(* IEC 61131-3 sources: volt/packages/volt-lsp-iec/test-corpus/lenze-mid/Device/Plc Logic/Application/Library Manager/L_OEEA_BaseDependency, 3.26.4.8 (Lenze), 88 files *)

(* ---- ENUMOEECALCULATIONMODE.dut ---- *)
TYPE ENUMOEECALCULATIONMODE :
(
	STANDARD := 0,
	PART_SUMMERY := 1
);
END_TYPE

(* ---- ENUMOEEPARTTARGETMODE.dut ---- *)
TYPE ENUMOEEPARTTARGETMODE :
(
	SHIFTPARTTARGET := 0,
	PRODUCTPARTTARGET := 1
);
END_TYPE

(* ---- ENUMRUNRATEFREQUENCE.dut ---- *)
TYPE ENUMRUNRATEFREQUENCE :
(
	HOUR_1X := 1,
	HOUR_2X := 2,
	HOUR_4X := 4
);
END_TYPE

(* ---- ENUMSHIFTMODE.dut ---- *)
TYPE ENUMSHIFTMODE :
(
	SHIFT := 0,
	HOURS24 := 1,
	NOSCHEDULE := 2,
	SHIFT7DAYS := 3,
	HOURS24_7DAYS := 4
);
END_TYPE

(* ---- RT_DOWNTIME.dut ---- *)
TYPE RT_DOWNTIME :
STRUCT
	PARA : ARRAY [0..19] OF sc_RT_Downtime;
END_STRUCT
END_TYPE

(* ---- RT_STATUS_STRUCT.dut ---- *)
TYPE RT_STATUS_STRUCT :
STRUCT
	STATIONID : DINT;
	PARTID : DINT;
	TOTALPARTSOK : DINT;
	TOTALPARTSNOK : DINT;
	TOTALPARTSOK_2 : DINT;
	TOTALPARTSNOK_2 : DINT;
	PARTTYPEID : DINT;
	PARTTYPESTR : STRING(100);
	PRODMODE : INT;
	PRODMODESTR : STRING;
	PARTCYCLETIME : REAL;
	OPCYCLETIME : REAL;
	ALIVECOUNTER : DINT;
	ERROR : BOOL;
	WARNING : BOOL;
	DOWNTIMECODE : INT;
	SDOWNTIMESTR : STRING;
	REASONCODE : DINT;
	REASONCODESTR : STRING;
	DOWNTIMEACTIVE : BOOL;
END_STRUCT
END_TYPE

(* ---- RT_TIMER.dut ---- *)
TYPE RT_TIMER :
STRUCT
	TOK_PART : TIME;
	TNOK_PART : TIME;
	TOK_PART2 : TIME;
	TNOK_PART2 : TIME;
	TALIVECOUNTER : TIME;
	TERROR : ARRAY [0..19] OF TIME;
	TERRORDURATION : ARRAY [0..19] OF TIME;
	TWARNING : TIME;
	TWARNINGDURATION : TIME;
	TPARTTYPECHANGE : TIME;
	TPARTCYCLETIME : TIME;
	TOPCYCLETIME : TIME;
END_STRUCT
END_TYPE

(* ---- SC_RT_DOWNTIME.dut ---- *)
TYPE SC_RT_DOWNTIME :
STRUCT
	PRODUCTIONMODE : INT;
	DOWNTIMECODE : INT;
	REASONCODE : DINT;
	SREASONCODESTR : STRING;
END_STRUCT
END_TYPE

(* ---- SCACCESSPOINTS.dut ---- *)
TYPE SCACCESSPOINTS :
STRUCT
	TACTUALPLANNEDPRODUCTION : TIME;
	TSHIFTPLANNEDPRODUCTION : TIME;
	TACTUALALLTIME : TIME;
	TACTUALRUNTIME : TIME;
	TDOWNTIME : TIME;
	TORGDOWNTIME : TIME;
	TNONPRODUCTIVETIME : TIME;
	DIACTUALALLTIME : DINT;
	DIACTUALPLANNEDPRODUCTION : DINT;
	DISHIFTPLANNEDPRODUCTION : DINT;
	DIACTUALRUNTIME : DINT;
	DIDOWNTIME : DINT;
	DIORGDOWNTIME : DINT;
	DINONPRODUCTIVETIME : DINT;
	LRPARTSUMMERY : LREAL;
	LRACTUALPARTCOUNT : LREAL;
	RINCONSISTENTPARTCOUNTDEVIATION : REAL;
	XPRODUCTIONTARGETREACHED : BOOL;
	XCHANGEOVERTIMEACTIVE : BOOL;
	XCHANGEOVERTIMEEXCEEDED : BOOL;
END_STRUCT
END_TYPE

(* ---- SCACTUALPRODUCTION.dut ---- *)
TYPE SCACTUALPRODUCTION :
STRUCT
	XPRODUCTIONACTIVE : BOOL;
	XPRODUCTIONHOLD : BOOL;
	EOEECALCMODE : enumOEECalculationMode;
	EOEEPARTTARGETMODE : enumOEEPartTargetMode;
	IOEEKPIDECIMALS : INT := 1;
	RSETSPEEDVALUE : REAL;
	RSETSPEEDPERCENT : REAL;
	ITRIGGER : INT;
END_STRUCT
END_TYPE

(* ---- SCBATCH.dut ---- *)
TYPE SCBATCH :
STRUCT
	DIID : DINT;
	DIJOBID : DINT;
	SJOBNO : STRING;
	DIJOBTARGET : DINT;
END_STRUCT
END_TYPE

(* ---- SCBATCHPRODUCTEND.dut ---- *)
TYPE SCBATCHPRODUCTEND :
STRUCT
	XONBATCHIDCHANGE : BOOL;
	XONPRODUCTIDCHANGE : BOOL;
	XONPRODUCTNAMECHANGE : BOOL;
	XONTECHNICALCYCLETIMECHANGE : BOOL;
	XONPOWERUPEVENT : BOOL;
	XONSHIFTENDEVENT : BOOL;
END_STRUCT
END_TYPE

(* ---- SCBREAKSCHEDULE.dut ---- *)
TYPE SCBREAKSCHEDULE :
STRUCT
	UISTARTHOUR : UINT;
	UISTARTMINUTE : UINT;
	UIENDHOUR : UINT;
	UIENDMINUTE : UINT;
	SBREAKNAME : STRING(uiShiftName);
	UISHIFTNO : UINT;
	XACTIVE : BOOL;
END_STRUCT
END_TYPE

(* ---- SCCLOUD.dut ---- *)
TYPE SCCLOUD :
STRUCT
	ISTATIONID : INT := 1;
	ROEERT : REAL;
	ROEETARGET : REAL;
	ROEECRUCIAL : REAL;
	RAVAILABILITY : REAL;
	RPERFORMANCE : REAL;
	RQUALITY : REAL;
	RTEEP : REAL;
	LRQUANTITYOK : LREAL;
	RQUANTITYTARGET : REAL;
	RPROGRESSIVETARGET : REAL;
	LRQUANTITYNOK : LREAL;
	LRACTUALTHROUGHPUT : LREAL;
	LRTARGETTHROUGHPUT : LREAL;
	RLASTCYCLETIME : REAL;
	RTECHNICALCYCLETIME : REAL;
	DINONPRODUCTIVETIME : DINT;
	DIDOWNTIME : DINT;
	DIORGDOWNTIME : DINT;
	DIACTUALPLANNEDPRODUCTION : DINT;
	DIACTUALRUNTIME : DINT;
	RSETSPEEDVALUE : REAL;
	RSETSPEEDPERCENT : REAL;
	ISHIFTID : INT;
	SSHIFT : STRING;
	SEVENT : STRING;
	IPRODUCTIONMODE : INT;
	SMODE : STRING;
	IDOWNTIMECATEGORY : INT;
	SDOWNTIMESTR : STRING;
	UDIDOWNTIMEREASON : UDINT;
	SREASONCODE : STRING;
	XCREATETICKET : BOOL;
	SCOMPONENTPATH : STRING;
	SSERIALNUMBER : STRING;
	ICALLFORSERVICE : INT;
	SSTARTTIME : STRING;
	SENDTIME : STRING;
	SSTARTBREAKTIME : STRING;
	SENDBREAKTIME : STRING;
	SSHIFTPLANNEDNONPRODUCTION : STRING;
	SSHIFTPLANNEDPRODUCTION : STRING;
	XACTIVE : BOOL;
	DIPARTID : DINT;
	SPARTTYPE : STRING;
	SUNITPRODUCT : STRING;
	SUNITSPEED : STRING;
	SDOWNTIME_WA_ER : STRING;
	SDATETIME : STRING;
	LRPARTCOUNT_RR : LREAL;
	LRQUANTITYOK_RR : LREAL;
	RINTERVALTARGET_RR : REAL;
	SDATETIME_RR : STRING;
	ITRIGGER_RR : INT;
	ITRIGGER_SETTINGS : INT;
END_STRUCT
END_TYPE

(* ---- SCCLOUDTICKETSYSTEM.dut ---- *)
TYPE SCCLOUDTICKETSYSTEM :
STRUCT
	IDOWNTIMECATEGORY : INT;
	SDOWNTIMESTR : STRING;
	UDIDOWNTIMEREASON : UDINT;
	SREASONCODE : STRING;
	XCREATETICKET : BOOL;
	SCOMPONENTPATH : STRING;
END_STRUCT
END_TYPE

(* ---- SCCURRENTSHIFTVALUES.dut ---- *)
TYPE SCCURRENTSHIFTVALUES :
STRUCT
	SSHIFT : STRING(uiShiftName);
	ESHIFTMODE : enumShiftMode;
	IBREAK : INT;
	SBREAK : STRING(uiShiftName);
	ESETWEEKDAY : RTCLK.WEEKDAY;
	DTSETWEEKSTARTTIME : TIME_OF_DAY;
	XSHIFTCHANGEEVENT : BOOL;
	XSHIFTCHANGESTOREEVENT : BOOL;
	XSCHEDULEDDOWNTIME : BOOL;
	TSHIFTPLANNEDNONPRODUCTION : TIME;
	XSHIFTDATAPROLONGED : BOOL;
	XSHIFTDAYSTARTPROLONGED : BOOL;
	XSHIFTDAYENDPROLONGED : BOOL;
	XPOWERONCYCLEPROLONGED : BOOL;
END_STRUCT
END_TYPE

(* ---- SCCURRENTSHIFTVALUES_BASE.dut ---- *)
TYPE SCCURRENTSHIFTVALUES_BASE :
STRUCT
	ISHIFT : INT;
	ISHIFTPREVIOUS : INT;
	XACTIVE : BOOL;
	EACTUALWEEKDAY : RTCLK.WEEKDAY;
	DTCURRENTTIME : TIME_OF_DAY;
	DTCURRENTDATE : DATE;
	DTSTARTTIME : TIME_OF_DAY;
	DTENDTIME : TIME_OF_DAY;
	TOFFSETSTARTTIME : TIME;
	DTSTARTBREAKTIME : TIME_OF_DAY;
	DTENDBREAKTIME : TIME_OF_DAY;
	DTDATEANDTIME : DATE_AND_TIME;
	DWCURRENTUTC_TIME : DWORD;
END_STRUCT
END_TYPE

(* ---- SCCUTAVERAGEREAL.dut ---- *)
TYPE SCCUTAVERAGEREAL :
STRUCT
	RREALINPUTVALUE : REAL;
	RINVALUE : REAL;
	SCUTREALSTR : STRING;
	RCUTREAL : REAL;
	LRCUTREAL : LREAL;
	IARRAYINDEX : INT;
	ARVALUEARRAY : ARRAY [0..60] OF REAL;
	RAVERAGEVALUE : REAL;
	RLASTREALVALUE : REAL;
END_STRUCT
END_TYPE

(* ---- SCDATEANDTIME.dut ---- *)
TYPE SCDATEANDTIME :
STRUCT
	UIYEAR : UINT;
	UIMONTH : UINT;
	UIDAY : UINT;
	UIHOUR : UINT;
	UIMINUTE : UINT;
	UISECOND : UINT;
END_STRUCT
END_TYPE

(* ---- SCDATETIMESTR.dut ---- *)
TYPE SCDATETIMESTR :
STRUCT
	SDATETIME : STRING;
	SSTARTTIME : STRING;
	SENDTIME : STRING;
	SSHIFTPLANNEDPRODUCTION : STRING;
	SSHIFTPLANNEDNONPRODUCTION : STRING;
	SSTARTBREAKTIME : STRING;
	SENDBREAKTIME : STRING;
END_STRUCT
END_TYPE

(* ---- SCDAYSCHEDULE.dut ---- *)
TYPE SCDAYSCHEDULE :
STRUCT
	ASCSHIFTSCHEDULE : ARRAY [1..uiNoOfShifts] OF scShiftSchedule;
	INUMBEROFSHIFTS : INT := UINT_TO_INT(uiNoOfShifts);
	ASCSBREAKSCHEDULE : ARRAY [1..uiNoOfBreaks] OF scBreakSchedule;
	INUMBEROFBREAKS : INT := UINT_TO_INT(uiNoOfBreaks);
END_STRUCT
END_TYPE

(* ---- SCDOWNTIME.dut ---- *)
TYPE SCDOWNTIME :
STRUCT
	SCPRODUCTIONMODES : ARRAY [0..uiNoOfProductionModes] OF scProductionModes;
	SCDOWNTIMECATEGORIES : ARRAY [0..uiNoOfDowntimeCategories] OF scDowntimeCategories;
	SCTOP3DOWNTIME : scVisuTop3Downtime;
	SCTOP3PRODUCTIONMODE : scVisuTop3ProductionMode;
	SCTOP3PERFORMANCELOSSES : scVisuTop3ProductionMode;
END_STRUCT
END_TYPE

(* ---- SCDOWNTIME_BASE.dut ---- *)
TYPE SCDOWNTIME_BASE :
STRUCT
	SDATETIME : STRING;
	SCLOGVALUES : ARRAY [0..uimaxLogSize] OF scDowntime_logValues;
	SRESULT : ARRAY [0..uimaxLogSize] OF STRING(255);
END_STRUCT
END_TYPE

(* ---- SCDOWNTIME_LOG.dut ---- *)
TYPE SCDOWNTIME_LOG :
STRUCT
	SRESULT : ARRAY [0..uimaxLogSize] OF STRING(255);
END_STRUCT
END_TYPE

(* ---- SCDOWNTIME_LOG_BASE.dut ---- *)
TYPE SCDOWNTIME_LOG_BASE :
STRUCT
	SCLOGVALUES : ARRAY [0..uimaxLogSize] OF scDowntime_logValues;
END_STRUCT
END_TYPE

(* ---- SCDOWNTIME_LOGVALUES.dut ---- *)
TYPE SCDOWNTIME_LOGVALUES :
STRUCT
	DTDATETIME : DATE_AND_TIME;
	IPRODUCTIONMODE : INT;
	IMODEBREAK : INT;
	IDOWNTIMECATEGORY : INT;
	UDIDOWNTIMEREASON : UDINT;
	DIRUNTIME : DINT;
	TDURATION : TIME;
END_STRUCT
END_TYPE

(* ---- SCDOWNTIMECATEGORIES.dut ---- *)
TYPE SCDOWNTIMECATEGORIES :
STRUCT
	IDOWNTIMECATEGORY : INT;
	SDOWNTIMESTR : STRING;
	XDOWNTIMEHISTORY : BOOL;
	XWARNING : BOOL;
	XERROR : BOOL;
	UIPRIORITY : UINT;
	DIDURATION : DINT;
	DIFREQUENCY : DINT;
	DIRUNTIME : DINT;
END_STRUCT
END_TYPE

(* ---- SCINTERNALDOWNVAR.dut ---- *)
TYPE SCINTERNALDOWNVAR :
STRUCT
	ILASTPRODUCTIONMODE : INT;
	ILASTDOWNTIMECATEGORY : INT := DINT_TO_INT(uiNoOfDowntimeCategories);
	UDILASTDOWNTIMEREASON : UDINT;
	ILOGINDEX : UINT;
	DTLASTDATETIME : DATE_AND_TIME;
END_STRUCT
END_TYPE

(* ---- SCINTERNALPRODUCTIONDATA.dut ---- *)
TYPE SCINTERNALPRODUCTIONDATA :
STRUCT
	RPARTTARGET : REAL;
	DTPRODUCTIONSTARTDATETIME : DATE_AND_TIME;
	DTPRODUCTIONENDDATETIME : DATE_AND_TIME;
	DTPRODUCTIONHOLDDATETIME : DATE_AND_TIME;
	DTSTARTTIME : TIME_OF_DAY;
	DTENDTIME : TIME_OF_DAY;
	DTSTARTBREAKTIME : TIME_OF_DAY;
	DTENDBREAKTIME : TIME_OF_DAY;
	TSHIFTPLANNEDNONPRODUCTION : TIME;
	IPREVIOUSRUN : INT;
	IACTUALRUN : INT;
END_STRUCT
END_TYPE

(* ---- SCINTERNALVAR.dut ---- *)
TYPE SCINTERNALVAR :
STRUCT
	SCPARTCOUNTER : scPartCounter;
	SCPARTCOUNTERDIFF : scPartCounter;
	RLASTMACHINECYCLETIME : REAL;
	LRPARTCOUNT : LREAL;
	RINTERVALTARGET : REAL;
	ISHFTCHANGECOUNTER : INT;
	LRLASTPARTSOK : LREAL;
	LRLASTPARTSNOK : LREAL;
	DILASTACTUALTIME : DINT;
	DIACTUALTIMEDIFF : DINT;
	SCAP : scAccessPoints;
	DTLASTDATETIME : DATE_AND_TIME;
	LRQUANTITYOK : LREAL;
	LRQUANTITYNOK : LREAL;
	SCPRODUCTTYPE : scProductCounts;
	SCSHIFTOEE : scShiftOEEStore;
	DILASTPLANNEDPRODUCTION : DINT;
	RLASTPARTTARGET : REAL;
END_STRUCT
END_TYPE

(* ---- SCMACHINEDATA.dut ---- *)
TYPE SCMACHINEDATA :
STRUCT
	SMODEBREAK : STRING;
	SCSHIFTDATA : scShiftData_base;
	SCPRODUCTDATA : scProduct;
	SCBUTTONS : scVisuButtons_base;
END_STRUCT
END_TYPE

(* ---- SCMACHINEDATA_BASE.dut ---- *)
TYPE SCMACHINEDATA_BASE :
STRUCT
	STATIONID : INT := 1;
	IPRODUCTIONMODE : INT;
	XDOWNTIMEACTIVE : BOOL;
	XORGDOWNTIMEACTIVE : BOOL;
	XSCHEDULEDDOWNTIMEACTIVE : BOOL;
	IDOWNTIMECATEGORY : INT;
	UDIDOWNTIMEREASON : UDINT;
	IMODEBREAK : INT;
	IMODEPRODUCTION : INT;
	DITYPEID : DINT;
	SCPARTDATA : scPartCounter;
	SCSHIFTTARGETS : scShiftTargetsInput;
	SCPRODUCTION : scActualProduction;
END_STRUCT
END_TYPE

(* ---- SCOEE_PD.dut ---- *)
TYPE SCOEE_PD :
STRUCT
	SCPERFORMANCE : scPerformance;
	SCDOWNTIME : scDowntime;
	SCSHIFTHISTORY : ARRAY [1..3] OF scPerformance;
	SCSHIFTDOWNTIMEHISTORY : ARRAY [1..3] OF scDowntime;
	SCPDINTERNAL : scInternalVar;
END_STRUCT
END_TYPE

(* ---- SCOEE_VISUPD.dut ---- *)
TYPE SCOEE_VISUPD :
STRUCT
	ASCVISU_OUT_SHIFTSCHEDULE : ARRAY [1..uiNoOfShifts] OF scShiftSchedule;
	ASCVISU_OUT_BREAKSCHEDULE : ARRAY [1..uiNoOfBreaks] OF scBreakSchedule;
	ASCVISU_OUT_SHIFTTARGETS : ARRAY [1..uiNoOfShifts] OF scShiftTargetsInput_base;
END_STRUCT
END_TYPE

(* ---- SCPARTCORRECTIONINPUT.dut ---- *)
TYPE SCPARTCORRECTIONINPUT :
STRUCT
	ICORRECTIONMODE : INT;
	LRCOUNTOK_CORRECTION : ARRAY [1..uiNoOfPartCounter] OF LREAL;
	LRCOUNTNOK_CORRECTION : ARRAY [1..uiNoOfPartCounter] OF LREAL;
END_STRUCT
END_TYPE

(* ---- SCPARTCOUNTER.dut ---- *)
TYPE SCPARTCOUNTER :
STRUCT
	SCPARTCORRECTIONINPUT : scPartCorrectionInput;
END_STRUCT
END_TYPE

(* ---- SCPARTCOUNTER_BASE.dut ---- *)
TYPE SCPARTCOUNTER_BASE :
STRUCT
	LRCOUNTOK : ARRAY [1..uiNoOfPartCounter] OF LREAL;
	LRCOUNTNOK : ARRAY [1..uiNoOfPartCounter] OF LREAL;
	RLASTCYCLETIME : REAL;
	XOVERFLOWCOUNT : BOOL;
END_STRUCT
END_TYPE

(* ---- SCPDSHIFTDATA.dut ---- *)
TYPE SCPDSHIFTDATA :
STRUCT
	DISHIFTDAYCOUNT : DINT;
	IPREVIOUSHIFTDAYINDEX : INT;
END_STRUCT
END_TYPE

(* ---- SCPERFORMANCE.dut ---- *)
TYPE SCPERFORMANCE :
STRUCT
	ICALLFORSERVICE : INT;
	ITRIGGER_SETTINGS : INT;
	SCTHROUGHPUT : scThroughput;
	SCSHIFTINTERVAL : scShiftInterval;
	SCSHIFTVALUES : scCurrentShiftValues;
	SCSHIFTTARGETS : scShiftTargetsInput;
	SCDATETIMESTR : scDateTimeStr;
	SCPRODUCTION : scActualProduction;
	SCPRODUCT : scProduct;
	SCAP : scAccessPoints;
	SCRR : scRunRate;
END_STRUCT
END_TYPE

(* ---- SCPERFORMANCE_BASE.dut ---- *)
TYPE SCPERFORMANCE_BASE :
STRUCT
	ISTATIONID : INT := 1;
	ISHIFT : INT;
	ROEERT : REAL;
	RTEEP : REAL;
	RAVAILABILITY : REAL;
	RPERFORMANCE : REAL;
	RQUALITY : REAL;
	LRQUANTITYOK : LREAL;
	RPROGRESSIVETARGET : REAL;
	LRQUANTITYNOK : LREAL;
	RLASTCYCLETIME : REAL;
	IPRODUCTIONMODE : INT;
	IDOWNTIMECATEGORY : INT;
	UDIDOWNTIMEREASON : UDINT;
	DITYPEID : DINT;
	XSTATECHANGEPROLONGED : BOOL;
	XOEEKPIPROLONGED : BOOL;
END_STRUCT
END_TYPE

(* ---- SCPRODUCT.dut ---- *)
TYPE SCPRODUCT :
STRUCT
	DIPARTID : DINT;
	DIBATCHID : DINT;
	SCBATCHPRODUCTEND : scBatchProductEnd;
	XBATCHIDACTIVE : BOOL;
	ITRIGGER : INT;
END_STRUCT
END_TYPE

(* ---- SCPRODUCT_BASE.dut ---- *)
TYPE SCPRODUCT_BASE :
STRUCT
	DITYPEID : DINT;
	RPRODUCTTARGET : REAL;
	RTECHNICALCYCLETIME : REAL;
	STYPENAME : STRING;
	IUNITPRODUCTID : INT := 1;
	SUNITPRODUCT : STRING;
	IUNITSPEEDID : INT := 1;
	SUNITSPEED : STRING;
	INOOFPARTSPERFIXTURE : INT;
	RCHANGEOVERTIME : REAL;
END_STRUCT
END_TYPE

(* ---- SCPRODUCTCOUNTS.dut ---- *)
TYPE SCPRODUCTCOUNTS :
STRUCT
	DIBATCHID : DINT;
	DITYPEID : DINT;
	STYPENAME : STRING;
	RTECHNICALCYCLETIME : REAL;
	ROEERT : REAL;
	RAVAILABILITY : REAL;
	RPERFORMANCE : REAL;
	RQUALITY : REAL;
	LRPRODUCTQUANTITYOK : LREAL;
	LRPRODUCTQUANTITYNOK : LREAL;
	DIACTUALRUNTIME : DINT;
	DIACTUALPLANNEDPRODUCTION : DINT;
	DIPRODUCTTOTALUNSCHEDULEDDOWNTIME : DINT;
	DWSTARTUTC_TIME : DWORD;
	DTSTARTDATEANDTIME : DATE_AND_TIME;
END_STRUCT
END_TYPE

(* ---- SCPRODUCTIONMODEPACKML.dut ---- *)
TYPE SCPRODUCTIONMODEPACKML :
STRUCT
	ASMODE : ARRAY [0..uiNoOfProductionModes] OF STRING := ['Undefined', 'Clearing', 'Stopped', 'Starting', 'Idle', 'Suspended', 'Execute', 'Stopping', 'Aborting', 'Aborted', 'Holding', 'Held', 'Unholding', 'Suspending', 'Unsuspending', 'Resetting', 'Completing', 'Complete', 'Reserved_1', 'Reserved_2', 'Break'];
END_STRUCT
END_TYPE

(* ---- SCPRODUCTIONMODES.dut ---- *)
TYPE SCPRODUCTIONMODES :
STRUCT
	IPRODUCTIONMODE : INT;
	SMODE : STRING;
	XDOWNTIME : BOOL;
	XORGDOWNTIME : BOOL;
	UIPRIORITY : UINT;
	DIDURATION : DINT;
	DIFREQUENCY : DINT;
	DIRUNTIME : DINT;
END_STRUCT
END_TYPE

(* ---- SCRUNRATE.dut ---- *)
TYPE SCRUNRATE :
STRUCT
	SDATETIME : STRING;
	LRPARTCOUNT : LREAL;
	LRQUANTITYOK : LREAL;
	RINTERVALTARGET : REAL;
	XRUNRATESAVED : BOOL;
	ITRIGGER : INT;
END_STRUCT
END_TYPE

(* ---- SCSHIFTDATA_BASE.dut ---- *)
TYPE SCSHIFTDATA_BASE :
STRUCT
	XFIRSTERRORACTIVE : BOOL;
	XISWARNINGINFO : BOOL;
	SINTERVAL : STRING;
	SDOWNTIMESTR : STRING;
	SREASONCODE : STRING;
	SMODECOLOURCODE : STRING(6);
	IPRODUCTIONEVENTMODE : INT;
END_STRUCT
END_TYPE

(* ---- SCSHIFTINTERVAL.dut ---- *)
TYPE SCSHIFTINTERVAL :
STRUCT
	SEVENT : STRING(255);
	SSHIFTOEEKPIS : STRING(255);
	SPRODUCTOEEKPIS : STRING(255);
	ITRIGGERSTATECOUNT : INT;
END_STRUCT
END_TYPE

(* ---- SCSHIFTINTERVAL_BASE.dut ---- *)
TYPE SCSHIFTINTERVAL_BASE :
STRUCT
	IPRODUCTIONMODE : INT;
	XDOWNTIMEACTIVE : BOOL;
	XORGDOWNTIMEACTIVE : BOOL;
	XSUSPENDEDACTIVE : BOOL;
	IDOWNTIMECATEGORY : INT;
	IDOWNTIMEREASON : INT;
	SCSHIFTTARGETS : scShiftTargetsInput;
	IMODEBREAK : INT;
	IMODEPRODUCTION : INT;
END_STRUCT
END_TYPE

(* ---- SCSHIFTOEEHISTORY_BASE.dut ---- *)
TYPE SCSHIFTOEEHISTORY_BASE :
STRUCT
	SDATETIME : STRING;
	ISHIFT : INT;
	ROEERT : REAL;
	RAVAILABILITY : REAL;
	RPERFORMANCE : REAL;
	RQUALITY : REAL;
	LRQUANTITYOK : LREAL;
END_STRUCT
END_TYPE

(* ---- SCSHIFTOEESTORE.dut ---- *)
TYPE SCSHIFTOEESTORE :
STRUCT
	ISHIFT : INT;
	SSHIFT : STRING(uiShiftName);
	ROEERT : REAL;
	RAVAILABILITY : REAL;
	RPERFORMANCE : REAL;
	RQUALITY : REAL;
	LRQUANTITYOK : LREAL;
	LRQUANTITYNOK : LREAL;
	DITOTALUNSCHEDULEDDOWNTIME : DINT;
	DWCURRENTUTC_TIME : DWORD;
	DWSTARTUTC_TIME : DWORD;
	DTDATEANDTIME : DATE_AND_TIME;
END_STRUCT
END_TYPE

(* ---- SCSHIFTSCHEDULE.dut ---- *)
TYPE SCSHIFTSCHEDULE :
STRUCT
	UISTARTHOUR : UINT;
	UISTARTMINUTE : UINT;
	UIENDHOUR : UINT;
	UIENDMINUTE : UINT;
	SSHIFTNAME : STRING(uiShiftName);
	UISHIFTNO : UINT;
	XACTIVE : BOOL;
	RPARTTARGET : REAL;
END_STRUCT
END_TYPE

(* ---- SCSHIFTTARGETSINPUT.dut ---- *)
TYPE SCSHIFTTARGETSINPUT :
STRUCT
	RPARTTARGET : REAL;
	RTECHNICALCYCLETIME : REAL;
END_STRUCT
END_TYPE

(* ---- SCSHIFTTARGETSINPUT_BASE.dut ---- *)
TYPE SCSHIFTTARGETSINPUT_BASE :
STRUCT
	ROEETARGET : REAL;
	ROEELOWERLIMIT : REAL;
	ROEECRUCIAL : REAL;
END_STRUCT
END_TYPE

(* ---- SCTHROUGHPUT.dut ---- *)
TYPE SCTHROUGHPUT :
STRUCT
	LRACTUALTHROUGHPUT_MIN : LREAL;
	LRTARGETTHROUGHPUT_MIN : LREAL;
	LRACTUALTHROUGHPUT_HR : LREAL;
	LRTARGETTHROUGHPUT_HR : LREAL;
	LRBESTSHIFTTHROUGHPUT_HR : LREAL;
	LRWORSESHIFTTHROUGHPUT_HR : LREAL;
END_STRUCT
END_TYPE

(* ---- SCTRIGGER.dut ---- *)
TYPE SCTRIGGER :
STRUCT
	ERRFREQ : enumRunRateFrequence := enumRunRateFrequence.hour_4x;
	TTRIGGER_SETTINGS : TIME := TIME#60m0s0ms;
END_STRUCT
END_TYPE

(* ---- SCTRIGGER_BASE.dut ---- *)
TYPE SCTRIGGER_BASE :
STRUCT
	TTRIGGER_DURATION : TIME := TIME#1s0ms;
	TTRIGGER_OEEKPI : TIME := TIME#1m0s0ms;
	TTRIGGER_POWERONDELAY : TIME := TIME#1m0s0ms;
END_STRUCT
END_TYPE

(* ---- SCVISUACTUALSHIFTTIMES.dut ---- *)
TYPE SCVISUACTUALSHIFTTIMES :
STRUCT
	TACTUALPLANNEDPRODUCTION : TIME;
	TACTUALRUNTIME : TIME;
	TDOWNTIME : TIME;
	TNONPRODUCTIVETIME : TIME;
	DIACTUALPLANNEDPRODUCTION : DINT;
	DIACTUALRUNTIME : DINT;
END_STRUCT
END_TYPE

(* ---- SCVISUBUTTONS.dut ---- *)
TYPE SCVISUBUTTONS :
STRUCT
	ISHIFTDAYNUMBER : INT;
	ISHIFTSAVESELECTION : INT;
	XSAVESHIFTDATA : BOOL;
END_STRUCT
END_TYPE

(* ---- SCVISUBUTTONS_BASE.dut ---- *)
TYPE SCVISUBUTTONS_BASE :
STRUCT
	XCALLFORSERVICE : BOOL;
END_STRUCT
END_TYPE

(* ---- SCVISUPERFORMANCEDASHBOARD.dut ---- *)
TYPE SCVISUPERFORMANCEDASHBOARD :
STRUCT
	SCSHIFTHISTORY : scVisuShiftHistory;
	SCACTUALSHIFTTIMES : scVisuActualShiftTimes;
	SCTOP3DOWNTIME : scVisuTop3Downtime;
	SCTOP3PRODUCTIONMODE : scVisuTop3ProductionMode;
	SCPRODUCTIONSTATUS : scVisuProductionStatus;
END_STRUCT
END_TYPE

(* ---- SCVISUPRODUCTIONSTATUS.dut ---- *)
TYPE SCVISUPRODUCTIONSTATUS :
STRUCT
	IUNITPRODUCTID : INT := 1;
	IUNITSPEEDID : INT := 1;
END_STRUCT
END_TYPE

(* ---- SCVISUPRODUCTIONSTATUS_BASE.dut ---- *)
TYPE SCVISUPRODUCTIONSTATUS_BASE :
STRUCT
	IPRODUCTIONSTATE : INT;
	TSTATERUNTIME : TIME;
	TSTATETOTALTIME : TIME;
	DISTATERUNTIME : DINT;
	DISTATETOTALTIME : DINT;
	DOWNTIME_WA_ER : STRING;
END_STRUCT
END_TYPE

(* ---- SCVISUSHIFTHISTORY.dut ---- *)
TYPE SCVISUSHIFTHISTORY :
STRUCT
	ISHIFT : ARRAY [0..(uiNoOfShifts - 1)] OF INT;
	SSHIFT : ARRAY [0..(uiNoOfShifts - 1)] OF STRING(uiShiftName);
	ROEERT : ARRAY [0..(uiNoOfShifts - 1)] OF REAL;
	LRQUANTITYOK : ARRAY [0..(uiNoOfShifts - 1)] OF LREAL;
END_STRUCT
END_TYPE

(* ---- SCVISUSHIFTHISTORY_BASE.dut ---- *)
TYPE SCVISUSHIFTHISTORY_BASE :
STRUCT
	SCSHIFTACTUAL_BASE : scShiftOEEHistory_base;
	SCSHIFTHISTORY : ARRAY [0..(uiNoOfShifts - 1)] OF scShiftOEEHistory_base;
END_STRUCT
END_TYPE

(* ---- SCVISUTHROUGHPUT.dut ---- *)
TYPE SCVISUTHROUGHPUT :
STRUCT
	LRBESTSHIFTTHROUGHPUT_HR : LREAL;
	LRWORSESHIFTTHROUGHPUT_HR : LREAL;
END_STRUCT
END_TYPE

(* ---- SCVISUTOP3DOWNTIME.dut ---- *)
TYPE SCVISUTOP3DOWNTIME :
STRUCT
	SCDOWNTIMECATEGORIES : ARRAY [0..2] OF scDowntimeCategories;
END_STRUCT
END_TYPE

(* ---- SCVISUTOP3PRODUCTIONMODE.dut ---- *)
TYPE SCVISUTOP3PRODUCTIONMODE :
STRUCT
	SCPRODUCTIONMODES : ARRAY [0..2] OF scProductionModes;
END_STRUCT
END_TYPE

(* ---- SCXAXIS_TREND.dut ---- *)
TYPE SCXAXIS_TREND :
STRUCT
	AXIS : ARRAY [0..imaxSizeXY_TREND] OF DATE_AND_TIME;
	AXIS2 : ARRAY [0..imaxSizeXY_TREND] OF DINT;
	AXIS3 : ARRAY [0..imaxSizeXY_TREND] OF INT;
END_STRUCT
END_TYPE

(* ---- SCYAXIS_TREND.dut ---- *)
TYPE SCYAXIS_TREND :
STRUCT
	AXIS_ACTUAL : ARRAY [0..GVL_Const_Production_log.imaxSizeXY_TREND] OF LREAL;
	AXIS_TARGET : ARRAY [0..GVL_Const_Production_log.imaxSizeXY_TREND] OF LREAL;
END_STRUCT
END_TYPE

(* ---- GVL_CONST_PRODUCTION_LOG.gvl ---- *)
VAR_GLOBAL
	IMAXSIZEXY_TREND : INT := 100;
END_VAR

(* ---- GVL_GLOBAL_CONSTANTS.gvl ---- *)
VAR_GLOBAL
	UIMAXLOGSIZE : UINT := 50;
	IMAXFIELDS : INT := 30;
END_VAR

(* ---- GVL_MPCONSTS.gvl ---- *)
VAR_GLOBAL
	UINOOFPARTCOUNTER : UINT := 2;
	UINOOFPRODUCTIONMODES : UINT := 20;
	UINOOFDOWNTIMECATEGORIES : UINT := 99;
END_VAR

(* ---- GVL_SSCONSTS.gvl ---- *)
VAR_GLOBAL
	UINOOFSHIFTS : UINT := 3;
	UIDAYSCHEDULE : UINT := 7;
	UISHIFTNAME : UINT := 80;
	UINOOFBREAKS : UINT := 9;
END_VAR

(* ---- VERSIONCONSTANTS.gvl ---- *)
VAR_GLOBAL
	GC_BYAMOUNTOFGENERALDATA : BYTE := 50;
	GC_BYAMOUNTDOWNTIMEERRORS : BYTE := 10;
	GC_IFILTERSAMPLES : INT := 20;
END_VAR

(* ---- BOOL_TO_SQLSTRING.pou ---- *)
FUNCTION BOOL_TO_SQLSTRING : STRING
VAR_INPUT
	XBOOLVALUE : BOOL;
END_VAR
END_FUNCTION

(* ---- CALC_UNIXTIME.pou ---- *)
FUNCTION CALC_UNIXTIME : DINT
VAR_INPUT
	DTACTUALDATETIME : DATE_AND_TIME;
END_VAR
END_FUNCTION

(* ---- CONVERTDATETIME_TO_STR.pou ---- *)
FUNCTION CONVERTDATETIME_TO_STR : STRING
VAR_INPUT
	DTTIME_VALUE : DATE_AND_TIME;
END_VAR
END_FUNCTION

(* ---- CONVERTTIME_TO_STR.pou ---- *)
FUNCTION CONVERTTIME_TO_STR : STRING
VAR_INPUT
	TTIME_VALUE : TIME;
END_VAR
END_FUNCTION

(* ---- CONVERTTOD_TO_STR.pou ---- *)
FUNCTION CONVERTTOD_TO_STR : STRING
VAR_INPUT
	TODTIME_VALUE : TIME_OF_DAY;
END_VAR
END_FUNCTION

(* ---- CUTDECIMALLREALVALUE.pou ---- *)
FUNCTION CUTDECIMALLREALVALUE : LREAL
VAR_INPUT
	LRVALUE : LREAL;
	INOOFDECIMAL : INT;
END_VAR
END_FUNCTION

(* ---- CUTDECIMALREALVALUE.pou ---- *)
FUNCTION CUTDECIMALREALVALUE : REAL
VAR_INPUT
	RVALUE : REAL;
	INOOFDECIMAL : INT;
END_VAR
END_FUNCTION

(* ---- CUTREALVALUE.pou ---- *)
FUNCTION CUTREALVALUE : REAL
VAR_INPUT
	RVALUE : REAL;
	INOOFDECIMAL : INT;
	INOOFAVERAGECOUNT : INT;
END_VAR
VAR_IN_OUT
	SCCUTAVERAGEREAL : scCutAverageReal;
END_VAR
END_FUNCTION

(* ---- STRING_TO_SQLSTRING.pou ---- *)
FUNCTION STRING_TO_SQLSTRING : STRING
VAR_INPUT
	SSTRINGVALUE : STRING;
END_VAR
END_FUNCTION

(* ---- TIMEPERIOD.pou ---- *)
FUNCTION TIMEPERIOD : TIME
VAR_INPUT
	DTSTARTTIME : TIME_OF_DAY;
	DTENDTIME : TIME_OF_DAY;
END_VAR
END_FUNCTION

(* ---- TOD_TO_SECONDS.pou ---- *)
FUNCTION TOD_TO_SECONDS : DINT
VAR_INPUT
	TODTIME : TIME_OF_DAY;
END_VAR
END_FUNCTION

(* ---- TODCONCAT_SECONDVALUE.pou ---- *)
FUNCTION TODCONCAT_SECONDVALUE : TIME_OF_DAY
VAR_INPUT
	DISECONDSVALUE : DINT;
END_VAR
END_FUNCTION

(* ---- TODSPLIT_DAYCHANGECALC.pou ---- *)
FUNCTION TODSPLIT_DAYCHANGECALC : DINT
VAR_INPUT
	TODTIMEHIGH : TIME_OF_DAY;
	TODTIMELOW : TIME_OF_DAY;
	PUIHOUR : UINT;
	PUIMINUTE : UINT;
	PUISECOND : UINT;
	PUIMILLISECOND : UINT;
END_VAR
END_FUNCTION
